FUNCTION F_DwordToBitReal_1 : REAL
VAR_INPUT
	dwIn : DWORD;
END_VAR
VAR
	pt : POINTER TO REAL;
END_VAR

pt := ADR(dwIn);
F_DwordToBitReal := pt^;

END_FUNCTION

(* stored: Version 1.1.0.1, ProductVersion 3.1.4024.15
   POU F_DwordToBitReal_1: Id {5f1cd5e6-ade9-4c5d-b7e2-2d055bef9650}, SpecialFunc None *)
